Fanuc KAREL source: KB00176.KL

PROGRAM KB00176
%NOLOCKGROUP
%ENVIRONMENT REGOPE
VAR
  P1: INTEGER
  P2: XYZWPR
  P3: INTEGER
BEGIN
  P1 = 1
  P2.X = 1.0
  P3 = 1
  SET_POS_REG(P1, P2, P3)
END KB00176
